FUNCTION F_OPC_LOCAL (* OPC-UA-ID fuer einen lokalen Knoten: opc_ua[ACTION;NODE] *)
  (* Standard: 61499-1; Description: Copyright (c) 2026 Meisterschulen am Ostbahnhof This program and the accompanying materials are made available under the terms of the Eclipse Public License 2.0 which is available at https://www.eclipse.org/legal/epl-2.0/ SPDX-License-Identifier: EPL-2.0 *)
  (* Version 1.0, 2026-10-17, Franz Höpfinger, Meisterschulen am Ostbahnhof, initial implementation *)
  PACKAGE MyLib_OPC;
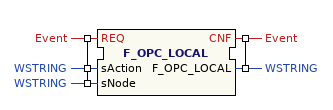
  EVENT_INPUT
    REQ WITH sAction, sNode;
  END_EVENT
  EVENT_OUTPUT
    CNF WITH F_OPC_LOCAL;
  END_EVENT
  VAR_INPUT
    sAction : WSTRING; (* ACTION, z.B. READ oder CREATE_METHOD *)
    sNode : WSTRING; (* Knoten, z.B. /Objects/X/Y,1:s=Y *)
  END_VAR
  VAR_OUTPUT
    F_OPC_LOCAL : WSTRING;
  END_VAR
  BODY IN ST:
PACKAGE MyLib_OPC;

(* OPC-UA-ID fuer einen lokalen Knoten: opc_ua[ACTION;NODE] *)
FUNCTION F_OPC_LOCAL : WSTRING

VAR_INPUT
	sAction : WSTRING; // ACTION, z.B. READ oder CREATE_METHOD
	sNode : WSTRING; // Knoten, z.B. /Objects/X/Y,1:s=Y
END_VAR

F_OPC_LOCAL := CONCAT("opc_ua[", sAction, ";", sNode, "]");

END_FUNCTION
  END_BODY
END_FUNCTION
